Fanuc KAREL source: kt00446.KL

-- PROVISIONAL review KL for V1013-1; original PC SHA256 623497cf41a629c7a82c3c50241ca8db61785963bb88cc6a9087745e85958422
-- Incomplete behavior may be omitted. Consult companion uncertainty JSON. Do not deploy.
PROGRAM KT00446
%NOLOCKGROUP
VAR
  S1 : STRING[80]
  S2 : STRING[80]
  OUT : BOOLEAN
BEGIN
  -- UNRESOLVED_PC offsets 5-14; opcodes 3F,75
  -- UNRESOLVED_PC offsets 19-28; opcodes 3F,75
  -- UNRESOLVED_PC offsets 33-42; opcodes 3F,75
  -- UNRESOLVED_PC offsets 47-56; opcodes 3F,75
  -- UNRESOLVED_PC offsets 61-80; opcodes 73,73,88,23
  -- UNRESOLVED_PC offsets 85-89; opcodes 7F
END KT00446
